Staubli VAL3: log.dtx

num nIndex = 14
num nLogType[300]
  [0] = 2
  [1] = 2
  [2] = 2
  [3] = 2
  [4] = 2
  [5] = 2
  [6] = 2
  [7] = 2
  [8] = 2
  [9] = 2
  [10] = 2
  [11] = 2
  [12] = 3
  [13] = 1
  [14] = 2
  [15] = 2
  [16] = 1
  [17] = 3
  [18] = 3
  [19] = 1
  [20] = 3
  [21] = 1
  [22] = 2
  [23] = 3
  [24] = 2
  [25] = 3
  [26] = 3
  [27] = 2
  [28] = 2
  [29] = 2
  [30] = 3
  [31] = 3
  [32] = 3
  [33] = 3
  [34] = 3
  [35] = 3
  [36] = 3
  [37] = 3
  [38] = 3
  [39] = 3
  [40] = 1
  [41] = 3
  [42] = 1
  [43] = 3
  [44] = 1
  [45] = 2
  [46] = 3
  [47] = 2
  [48] = 3
  [49] = 3
  [50] = 2
  [51] = 3
  [52] = 2
  [53] = 1
  [54] = 3
  [55] = 1
  [56] = 3
  [57] = 1
  [58] = 3
  [59] = 1
  [60] = 3
  [61] = 1
  [62] = 3
  [63] = 1
  [64] = 1
  [65] = 3
  [66] = 3
  [67] = 3
  [68] = 3
  [69] = 3
  [70] = 3
  [71] = 3
  [72] = 3
  [73] = 3
  [74] = 3
  [75] = 1
  [76] = 3
  [77] = 1
  [78] = 3
  [79] = 1
  [80] = 2
  [81] = 3
  [82] = 2
  [83] = 3
  [84] = 3
  [85] = 2
  [86] = 3
  [87] = 3
  [88] = 3
  [89] = 3
  [90] = 3
  [91] = 1
  [92] = 3
  [93] = 3
  [94] = 3
  [95] = 1
  [96] = 2
  [97] = 3
  [98] = 3
  [99] = 2
  [100] = 3
  [101] = 3
  [102] = 3
  [103] = 3
  [104] = 3
  [105] = 3
  [106] = 3
  [107] = 3
  [108] = 3
  [109] = 3
  [110] = 3
  [111] = 3
  [112] = 3
  [113] = 1
  [114] = 3
  [115] = 1
  [116] = 3
  [117] = 3
  [118] = 1
  [119] = 2
  [120] = 3
  [121] = 2
  [122] = 2
  [123] = 2
  [124] = 3
  [125] = 3
  [126] = 3
  [127] = 3
  [128] = 3
  [129] = 2
  [130] = 3
  [131] = 2
  [132] = 3
  [133] = 2
  [134] = 3
  [135] = 2
  [136] = 3
  [137] = 2
  [138] = 3
  [139] = 2
  [140] = 3
  [141] = 2
  [142] = 3
  [143] = 3
  [144] = 2
  [145] = 2
  [146] = 2
  [147] = 2
  [148] = 2
  [149] = 2
  [150] = 2
  [151] = 2
  [152] = 2
  [153] = 2
  [154] = 2
  [155] = 2
  [156] = 2
  [157] = 2
  [158] = 2
  [159] = 2
  [160] = 2
  [161] = 2
  [162] = 2
  [163] = 2
  [164] = 2
  [165] = 2
  [166] = 2
  [167] = 2
  [168] = 2
  [169] = 2
  [170] = 2
  [171] = 2
  [172] = 2
  [173] = 2
  [174] = 2
  [175] = 2
  [176] = 2
  [177] = 2
  [178] = 2
  [179] = 2
  [180] = 1
  [181] = 3
  [182] = 3
  [183] = 3
  [184] = 1
  [185] = 3
  [186] = 3
  [187] = 1
  [188] = 3
  [189] = 2
  [190] = 3
  [191] = 3
  [192] = 3
  [193] = 3
  [194] = 3
  [195] = 2
  [196] = 3
  [197] = 3
  [198] = 3
  [199] = 3
  [200] = 3
  [201] = 3
  [202] = 1
  [203] = 3
  [204] = 3
  [205] = 3
  [206] = 3
  [207] = 1
  [208] = 3
  [209] = 3
  [210] = 1
  [211] = 2
  [212] = 3
  [213] = 2
  [214] = 2
  [215] = 2
  [216] = 3
  [217] = 3
  [218] = 2
  [219] = 2
  [220] = 3
  [221] = 3
  [222] = 2
  [223] = 2
  [224] = 3
  [225] = 2
  [226] = 3
  [227] = 2
  [228] = 3
  [229] = 2
  [230] = 3
  [231] = 3
  [232] = 2
  [233] = 2
  [234] = 2
  [235] = 2
  [236] = 2
  [237] = 2
  [238] = 2
  [239] = 2
  [240] = 2
  [241] = 2
  [242] = 2
  [243] = 2
  [244] = 2
  [245] = 2
  [246] = 2
  [247] = 2
  [248] = 2
  [249] = 2
  [250] = 1
  [251] = 3
  [252] = 3
  [253] = 3
  [254] = 1
  [255] = 3
  [256] = 3
  [257] = 3
  [258] = 1
  [259] = 2
  [260] = 3
  [261] = 3
  [262] = 3
  [263] = 2
  [264] = 3
  [265] = 3
  [266] = 1
  [267] = 3
  [268] = 3
  [269] = 1
  [270] = 3
  [271] = 1
  [272] = 2
  [273] = 3
  [274] = 2
  [275] = 2
  [276] = 3
  [277] = 2
  [278] = 2
  [279] = 3
  [280] = 2
  [281] = 2
  [282] = 3
  [283] = 2
  [284] = 3
  [285] = 2
  [286] = 3
  [287] = 2
  [288] = 3
  [289] = 2
  [290] = 3
  [291] = 3
  [292] = 2
  [293] = 2
  [294] = 2
  [295] = 2
  [296] = 2
  [297] = 2
  [298] = 2
  [299] = 2
string sLog[300]
  [0] = "258.828 [路径信息]:移动到:12, L[271,-458,568,-7,-3,28]_spd=100%_b=50 09-16 10:48:04"
  [1] = "258.944 [路径信息]:移动到:13, L[271,-423,568,-7,-3,28]_spd=100%_b=50 09-16 10:48:04"
  [2] = "259.064 [路径信息]:移动到:14, L[241,-401,568,-7,-3,28]_spd=100%_b=50 09-16 10:48:05"
  [3] = "259.184 [路径信息]:移动到:15, L[189,-422,568,-7,-3,28]_spd=100%_b=50 09-16 10:48:05"
  [4] = "259.328 [路径信息]:移动到:16, L[189,-458,568,-7,-3,28]_spd=100%_b=50 09-16 10:48:05"
  [5] = "259.444 [路径信息]:移动到:17, L[159,-434,568,-7,-3,28]_spd=100%_b=50 09-16 10:48:05"
  [6] = "259.564 [路径信息]:移动到:18, L[121,-459,568,-7,-3,28]_spd=100%_b=50 09-16 10:48:06"
  [7] = "259.684 [路径信息]:移动到:19, L[121,-424,568,-7,-3,28]_spd=100%_b=50 09-16 10:48:06"
  [8] = "259.804 [路径信息]:移动到:20, L[90,-399,568,-7,-3,28]_spd=100%_b=50 09-16 10:48:06"
  [9] = "259.944 [路径信息]:移动到:21, L[40,-417,568,-7,-3,28]_spd=100%_b=50 09-16 10:48:06"
  [10] = "260.092 [路径信息]:移动到:22, L[40,-456,568,-7,-3,28]_spd=100%_b=50 09-16 10:48:07"
  [11] = "260.184 [路径信息]:移动到:23, L[3,-425,568,-7,-3,28]_spd=100%_b=50 09-16 10:48:07"
  [12] = "260.184 [信号信息]:dOut6=OFF 09-16 10:48:07"
  [13] = "261.184 [状态信息]:错误：-303. :0自动运行过程中伺服异常下电 09-16 10:48:09"
  [14] = "1112.913 [路径信息]:移动到:2, DOUT[70]-备用=TRUE 07-21 20:12:43"
  [15] = "1112.94  [路径信息]:移动到:3, wait->DIN[70]-备用=TRUE 07-21 20:12:43"
  [16] = "1294.838 [状态信息]:页面设置复位信号 07-21 20:17:28"
  [17] = "1297.928 [信号信息]:dOut10=OFF 07-21 20:17:33"
  [18] = "1298.8   [信号信息]:dOut6=ON 07-21 20:17:35"
  [19] = "1299.434 [状态信息]:程序号:1,J1MaxForce：0   ,J2MaxForce：152.6 ,J3MaxForce：73   ,J4MaxForce：1.3 ,J5MaxForce：10.03,J6MaxForce：0    07-21 20:17:36"
  [20] = "1299.434 [信号信息]:dOut1=ON 07-21 20:17:36"
  [21] = "1306.503 [状态信息]:当前处于生产状态 07-21 20:17:47"
  [22] = "1306.503 [路径信息]:移动到:0, DELAY = 1     s 07-21 20:17:47"
  [23] = "1306.503 [信号信息]:dOut2=ON 07-21 20:17:47"
  [24] = "1307.526 [路径信息]:移动到:1, L[1169,127,-142,15,129,-19]_spd=100%_b=0 07-21 20:17:48"
  [25] = "1307.526 [信号信息]:dOut8=ON 07-21 20:17:48"
  [26] = "1309.081 [信号信息]:dOut5=OFF 07-21 20:17:51"
  [27] = "1311.831 [路径信息]:移动到:2, L[1169,266,-142,15,129,-19]_spd=100%_b=0 07-21 20:17:55"
  [28] = "1316.763 [路径信息]:移动到轨迹PR01Washing001:3, WASH_DELAY = 0     s 07-21 20:18:03"
  [29] = "1316.784 [路径信息]:移动到:4, L[1169,266,-142,26,129,-19]_spd=100%_b=0 07-21 20:18:03"
  [30] = "1321.135 [信号信息]:dOut6=OFF 07-21 20:18:10"
  [31] = "180.317 [信号信息]:dOut97=ON 07-21 20:48:43"
  [32] = "196.059 [信号信息]:dOut6=ON 07-21 20:49:08"
  [33] = "196.677 [信号信息]:dOut8=ON 07-21 20:49:09"
  [34] = "197.418 [信号信息]:dOut97=OFF 07-21 20:49:10"
  [35] = "198.018 [信号信息]:dOut8=OFF 07-21 20:49:11"
  [36] = "199.801 [信号信息]:dOut8=ON 07-21 20:49:14"
  [37] = "203.867 [信号信息]:dOut5=ON 07-21 20:49:20"
  [38] = "204.256 [信号信息]:dOut8=OFF 07-21 20:49:21"
  [39] = "208.562 [信号信息]:dOut10=OFF 07-21 20:49:28"
  [40] = "212.136 [状态信息]:页面设置复位信号 07-21 20:49:33"
  [41] = "213.265 [信号信息]:dOut6=ON 07-21 20:49:35"
  [42] = "213.865 [状态信息]:当前处于ready状态 07-21 20:49:36"
  [43] = "213.887 [信号信息]:dOut1=ON 07-21 20:49:36"
  [44] = "251.032 [状态信息]:当前处于生产状态 07-21 20:50:34"
  [45] = "251.032 [路径信息]:移动到:0, DELAY = 1     s 07-21 20:50:34"
  [46] = "251.032 [信号信息]:dOut2=ON 07-21 20:50:34"
  [47] = "252.064 [路径信息]:移动到:1, L[1169,127,-142,15,129,-19]_spd=100%_b=0 07-21 20:50:36"
  [48] = "252.064 [信号信息]:dOut8=ON 07-21 20:50:36"
  [49] = "253.63  [信号信息]:dOut5=OFF 07-21 20:50:38"
  [50] = "256.347 [路径信息]:移动到:2, L[1169,266,-142,15,129,-19]_spd=100%_b=0 07-21 20:50:42"
  [51] = "261.222 [信号信息]:dOut6=OFF 07-21 20:50:50"
  [52] = "261.284 [路径信息]:移动到:4, L[1169,266,-142,26,129,-19]_spd=100%_b=0 07-21 20:50:50"
  [53] = "262.212 [状态信息]:错误：-303. :0自动运行过程中伺服异常下电 07-21 20:50:52"
  [54] = "262.733 [信号信息]:dOut11=ON 07-21 20:50:52"
  [55] = "262.759 [状态信息]:当前处于暂停状态 07-21 20:50:52"
  [56] = "262.759 [信号信息]:dOut3=ON 07-21 20:50:52"
  [57] = "264.227 [状态信息]:当前处于生产停止状态 07-21 20:50:55"
  [58] = "264.227 [信号信息]:dOut0=ON 07-21 20:50:55"
  [59] = "269.89  [状态信息]:收到页面点击清除报错! 07-21 20:51:04"
  [60] = "269.915 [信号信息]:dOut11=OFF 07-21 20:51:04"
  [61] = "273.022 [状态信息]:收到页面手动路径回Home点信号 07-21 20:51:09"
  [62] = "276.855 [信号信息]:dOut6=ON 07-21 20:51:15"
  [63] = "299.325 [状态信息]:页面设置复位信号 07-21 20:51:50"
  [64] = "301.959 [状态信息]:收到页面手动路径回Home点信号 07-21 20:51:54"
  [65] = "565.227 [信号信息]:dOut8=ON 07-21 20:58:47"
  [66] = "567.33  [信号信息]:dOut8=OFF 07-21 20:58:50"
  [67] = "571.862 [信号信息]:dOut8=ON 07-21 20:58:57"
  [68] = "572.394 [信号信息]:dOut8=OFF 07-21 20:58:58"
  [69] = "572.469 [信号信息]:dOut8=ON 07-21 20:58:58"
  [70] = "573.584 [信号信息]:dOut8=OFF 07-21 20:59:00"
  [71] = "575.243 [信号信息]:dOut8=ON 07-21 20:59:02"
  [72] = "575.802 [信号信息]:dOut5=ON 07-21 20:59:03"
  [73] = "576.029 [信号信息]:dOut8=OFF 07-21 20:59:04"
  [74] = "589.435 [信号信息]:dOut10=OFF 07-21 20:59:25"
  [75] = "604.459 [状态信息]:页面设置复位信号 07-21 20:59:48"
  [76] = "605.601 [信号信息]:dOut6=ON 07-21 20:59:50"
  [77] = "606.232 [状态信息]:程序号:1,J1MaxForce：67.45,J2MaxForce：264.18,J3MaxForce：102.39,J4MaxForce：8.71,J5MaxForce：19.2 ,J6MaxForce：1.88 07-21 20:59:51"
  [78] = "606.232 [信号信息]:dOut1=ON 07-21 20:59:51"
  [79] = "612.58  [状态信息]:当前处于生产状态 07-21 21:00:01"
  [80] = "612.58  [路径信息]:移动到:0, DELAY = 1     s 07-21 21:00:01"
  [81] = "612.58  [信号信息]:dOut2=ON 07-21 21:00:01"
  [82] = "613.621 [路径信息]:移动到:1, L[1169,127,-142,15,129,-19]_spd=100%_b=0 07-21 21:00:02"
  [83] = "613.621 [信号信息]:dOut8=ON 07-21 21:00:02"
  [84] = "615.161 [信号信息]:dOut5=OFF 07-21 21:00:05"
  [85] = "617.895 [路径信息]:移动到:2, L[1169,266,-142,15,129,-19]_spd=100%_b=0 07-21 21:00:09"
  [86] = "620.296 [信号信息]:dOut8=OFF 07-21 21:00:13"
  [87] = "620.788 [信号信息]:dOut6=OFF 07-21 21:00:14"
  [88] = "9.52  [信号信息]:dOut10=ON 09-16 10:39:57"
  [89] = "19.528 [信号信息]:dOut10=OFF 09-16 10:40:17"
  [90] = "60.184 [信号信息]:dIn0=ON 09-16 10:41:36"
  [91] = "60.312 [状态信息]:收到PLC复位信号 09-16 10:41:37"
  [92] = "60.828 [信号信息]:dIn0=OFF 09-16 10:41:38"
  [93] = "61.828 [信号信息]:dOut6=ON 09-16 10:41:40"
  [94] = "67.68  [信号信息]:dIn9=ON 09-16 10:41:51"
  [95] = "67.704 [状态信息]:收到PLC直接回Home点信号 09-16 10:41:51"
  [96] = "67.704 [路径信息]:直接回原点过程中 09-16 10:41:51"
  [97] = "67.704 [信号信息]:dOut8=ON 09-16 10:41:51"
  [98] = "68.564 [信号信息]:dOut5=ON 09-16 10:41:53"
  [99] = "68.796 [路径信息]:直接回原点完成 09-16 10:41:53"
  [100] = "68.796 [信号信息]:dOut6=OFF 09-16 10:41:53"
  [101] = "68.844 [信号信息]:dOut8=OFF 09-16 10:41:53"
  [102] = "69.076 [信号信息]:dOut0=ON 09-16 10:41:54"
  [103] = "69.404 [信号信息]:dIn9=OFF 09-16 10:41:54"
  [104] = "73.4   [信号信息]:dIn1=ON 09-16 10:42:02"
  [105] = "74.62  [信号信息]:dIn1=OFF 09-16 10:42:05"
  [106] = "87.112 [信号信息]:dOut8=ON 09-16 10:42:29"
  [107] = "87.18  [信号信息]:dOut8=OFF 09-16 10:42:29"
  [108] = "88.984 [信号信息]:dIn1=ON 09-16 10:42:33"
  [109] = "89.924 [信号信息]:dIn1=OFF 09-16 10:42:34"
  [110] = "102.18  [信号信息]:dIn1=ON 09-16 10:42:58"
  [111] = "109.252 [信号信息]:dIn1=OFF 09-16 10:43:12"
  [112] = "110.004 [信号信息]:dIn0=ON 09-16 10:43:14"
  [113] = "110.132 [状态信息]:收到PLC复位信号 09-16 10:43:14"
  [114] = "111.18  [信号信息]:dIn0=OFF 09-16 10:43:16"
  [115] = "112.78  [状态信息]:当前处于ready状态 09-16 10:43:19"
  [116] = "112.78  [信号信息]:dOut1=ON 09-16 10:43:19"
  [117] = "113.112 [信号信息]:dIn1=ON 09-16 10:43:20"
  [118] = "113.24  [状态信息]:当前处于生产状态 09-16 10:43:20"
  [119] = "113.24  [路径信息]:移动到:4, AOUT[4]-备用=0     09-16 10:43:20"
  [120] = "113.24  [信号信息]:dOut2=ON 09-16 10:43:20"
  [121] = "113.264 [路径信息]:移动到:10, DOUT[43]-吹干阀1=FALSE 09-16 10:43:20"
  [122] = "113.284 [路径信息]:移动到:14, DOUT[51]-吹干工作完成=FALSE 09-16 10:43:20"
  [123] = "113.308 [路径信息]:移动到:1, wait->DIN[20]-工作允许=TRUE 09-16 10:43:20"
  [124] = "114.424 [信号信息]:dIn1=OFF 09-16 10:43:22"
  [125] = "121.784 [信号信息]:dIn21=ON 09-16 10:43:37"
  [126] = "122.6   [信号信息]:dIn21=OFF 09-16 10:43:38"
  [127] = "125.18  [信号信息]:dIn40=ON 09-16 10:43:43"
  [128] = "125.82  [信号信息]:dIn40=OFF 09-16 10:43:45"
  [129] = "136.164 [路径信息]:移动到:0, DOUT[5]-机械人在home点=TRUE 09-16 10:44:05"
  [130] = "136.164 [信号信息]:dIn20=ON 09-16 10:44:05"
  [131] = "136.188 [路径信息]:移动到:2, DELAY = 0.5   s 09-16 10:44:05"
  [132] = "136.188 [信号信息]:dOut40=ON 09-16 10:44:05"
  [133] = "136.7   [路径信息]:移动到:3, wait->DIN[40]-私服位置到达=TRUE 09-16 10:44:06"
  [134] = "137.044 [信号信息]:dIn20=OFF 09-16 10:44:06"
  [135] = "138.724 [路径信息]:移动到:4, DELAY = 0.5   s 09-16 10:44:10"
  [136] = "138.724 [信号信息]:dIn40=ON 09-16 10:44:10"
  [137] = "139.232 [路径信息]:移动到:5, DOUT[40]-伺服旋转命令=FALSE 09-16 10:44:11"
  [138] = "139.232 [信号信息]:dOut40=OFF 09-16 10:44:11"
  [139] = "139.252 [路径信息]:移动到:2, L[61,-652,350,-2,-2,28]_spd=100%_b=50 09-16 10:44:11"
  [140] = "139.252 [信号信息]:dOut8=ON 09-16 10:44:11"
  [141] = "139.276 [路径信息]:移动到:3, L[489,-419,568,-7,-3,28]_spd=100%_b=50 09-16 10:44:11"
  [142] = "139.42  [信号信息]:dOut5=OFF 09-16 10:44:11"
  [143] = "139.744 [信号信息]:dIn40=OFF 09-16 10:44:12"
  [144] = "139.788 [路径信息]:移动到:4, L[489,-457,568,-7,-3,28]_spd=100%_b=50 09-16 10:44:12"
  [145] = "139.884 [路径信息]:移动到:5, L[459,-434,568,-7,-3,28]_spd=100%_b=50 09-16 10:44:12"
  [146] = "140.02  [路径信息]:移动到:6, L[427,-421,568,-7,-3,28]_spd=100%_b=50 09-16 10:44:12"
  [147] = "140.14  [路径信息]:移动到:7, L[427,-458,568,-7,-3,28]_spd=100%_b=50 09-16 10:44:12"
  [148] = "140.252 [路径信息]:移动到:8, L[393,-403,568,-7,-3,28]_spd=100%_b=50 09-16 10:44:13"
  [149] = "140.42  [路径信息]:移动到:9, L[345,-458,568,-7,-3,28]_spd=100%_b=50 09-16 10:44:13"
  [150] = "140.532 [路径信息]:移动到:10, L[345,-422,568,-7,-3,28]_spd=100%_b=50 09-16 10:44:13"
  [151] = "140.676 [路径信息]:移动到:11, L[312,-431,568,-7,-3,28]_spd=100%_b=50 09-16 10:44:14"
  [152] = "140.788 [路径信息]:移动到:12, L[271,-458,568,-7,-3,28]_spd=100%_b=50 09-16 10:44:14"
  [153] = "140.908 [路径信息]:移动到:13, L[271,-423,568,-7,-3,28]_spd=100%_b=50 09-16 10:44:14"
  [154] = "141.02  [路径信息]:移动到:14, L[241,-401,568,-7,-3,28]_spd=100%_b=50 09-16 10:44:14"
  [155] = "141.164 [路径信息]:移动到:15, L[189,-422,568,-7,-3,28]_spd=100%_b=50 09-16 10:44:14"
  [156] = "141.3   [路径信息]:移动到:16, L[189,-458,568,-7,-3,28]_spd=100%_b=50 09-16 10:44:15"
  [157] = "141.396 [路径信息]:移动到:17, L[159,-434,568,-7,-3,28]_spd=100%_b=50 09-16 10:44:15"
  [158] = "141.532 [路径信息]:移动到:18, L[121,-459,568,-7,-3,28]_spd=100%_b=50 09-16 10:44:15"
  [159] = "141.652 [路径信息]:移动到:19, L[121,-424,568,-7,-3,28]_spd=100%_b=50 09-16 10:44:15"
  [160] = "141.768 [路径信息]:移动到:20, L[90,-399,568,-7,-3,28]_spd=100%_b=50 09-16 10:44:16"
  [161] = "141.908 [路径信息]:移动到:21, L[40,-417,568,-7,-3,28]_spd=100%_b=50 09-16 10:44:16"
  [162] = "142.044 [路径信息]:移动到:22, L[40,-456,568,-7,-3,28]_spd=100%_b=50 09-16 10:44:16"
  [163] = "142.14  [路径信息]:移动到:23, L[3,-425,568,-7,-3,28]_spd=100%_b=50 09-16 10:44:16"
  [164] = "142.276 [路径信息]:移动到:24, L[-30,-459,568,-7,-3,28]_spd=100%_b=50 09-16 10:44:17"
  [165] = "142.396 [路径信息]:移动到:25, L[-30,-424,568,-7,-3,28]_spd=100%_b=50 09-16 10:44:17"
  [166] = "142.532 [路径信息]:移动到:26, L[-63,-402,568,-7,-3,28]_spd=100%_b=50 09-16 10:44:17"
  [167] = "142.652 [路径信息]:移动到:27, L[-112,-422,568,-7,-3,28]_spd=100%_b=50 09-16 10:44:17"
  [168] = "142.788 [路径信息]:移动到:28, L[-112,-459,568,-7,-3,28]_spd=100%_b=50 09-16 10:44:18"
  [169] = "142.908 [路径信息]:移动到:29, L[-149,-435,568,-7,-3,28]_spd=100%_b=50 09-16 10:44:18"
  [170] = "143.024 [路径信息]:移动到:30, L[-182,-460,568,-7,-3,28]_spd=100%_b=50 09-16 10:44:18"
  [171] = "143.14  [路径信息]:移动到:31, L[-182,-422,568,-7,-3,28]_spd=100%_b=50 09-16 10:44:18"
  [172] = "143.276 [路径信息]:移动到:32, L[-219,-406,568,-7,-3,28]_spd=100%_b=50 09-16 10:44:19"
  [173] = "143.42  [路径信息]:移动到:33, L[-267,-419,568,-7,-3,28]_spd=100%_b=50 09-16 10:44:19"
  [174] = "143.532 [路径信息]:移动到:34, L[-267,-457,568,-7,-3,28]_spd=100%_b=50 09-16 10:44:19"
  [175] = "143.676 [路径信息]:移动到:35, L[-308,-435,568,-7,-3,28]_spd=100%_b=50 09-16 10:44:19"
  [176] = "143.788 [路径信息]:移动到:36, L[-339,-459,568,-7,-3,28]_spd=100%_b=50 09-16 10:44:20"
  [177] = "143.908 [路径信息]:移动到:37, L[-339,-419,568,-7,-3,28]_spd=100%_b=50 09-16 10:44:20"
  [178] = "144.068 [路径信息]:移动到:38, L[-376,-400,568,-7,-3,28]_spd=100%_b=50 09-16 10:44:20"
  [179] = "144.164 [路径信息]:移动到:39, L[-338,-600,568,-7,-3,28]_spd=100%_b=50 09-16 10:44:20"
  [180] = "144.324 [状态信息]:页面设置停止信号 09-16 10:44:21"
  [181] = "144.324 [信号信息]:dOut2=OFF 09-16 10:44:21"
  [182] = "144.488 [信号信息]:dOut6=OFF 09-16 10:44:21"
  [183] = "144.556 [信号信息]:dOut8=OFF 09-16 10:44:21"
  [184] = "144.764 [状态信息]:当前处于生产停止状态 09-16 10:44:22"
  [185] = "144.764 [信号信息]:dOut42=OFF 09-16 10:44:22"
  [186] = "146.42  [信号信息]:dOut10=ON 09-16 10:44:25"
  [187] = "148.444 [状态信息]:收到页面手动路径回Home点信号 09-16 10:44:29"
  [188] = "150.532 [信号信息]:dOut6=ON 09-16 10:44:33"
  [189] = "151.724 [路径信息]:路径回原点过程中 09-16 10:44:35"
  [190] = "151.724 [信号信息]:dOut0=OFF 09-16 10:44:35"
  [191] = "154.7   [信号信息]:dOut8=ON 09-16 10:44:41"
  [192] = "179.3   [信号信息]:dOut8=OFF 09-16 10:45:29"
  [193] = "181.628 [信号信息]:dOut8=ON 09-16 10:45:33"
  [194] = "184.512 [信号信息]:dOut5=ON 09-16 10:45:39"
  [195] = "185.02  [路径信息]:路径回原点完成 09-16 10:45:40"
  [196] = "185.02  [信号信息]:dOut6=OFF 09-16 10:45:40"
  [197] = "185.3   [信号信息]:dOut0=ON 09-16 10:45:41"
  [198] = "188.236 [信号信息]:dOut10=OFF 09-16 10:45:46"
  [199] = "193.532 [信号信息]:dIn1=ON 09-16 10:45:57"
  [200] = "194.908 [信号信息]:dIn1=OFF 09-16 10:45:59"
  [201] = "195.468 [信号信息]:dIn0=ON 09-16 10:46:00"
  [202] = "195.596 [状态信息]:收到PLC复位信号 09-16 10:46:01"
  [203] = "196.128 [信号信息]:dIn0=OFF 09-16 10:46:02"
  [204] = "196.456 [信号信息]:dIn1=ON 09-16 10:46:02"
  [205] = "197.128 [信号信息]:dOut6=ON 09-16 10:46:04"
  [206] = "197.48  [信号信息]:dIn1=OFF 09-16 10:46:04"
  [207] = "197.74  [状态信息]:当前处于ready状态 09-16 10:46:05"
  [208] = "197.74  [信号信息]:dOut1=ON 09-16 10:46:05"
  [209] = "205.512 [信号信息]:dIn1=ON 09-16 10:46:20"
  [210] = "205.64  [状态信息]:当前处于生产状态 09-16 10:46:20"
  [211] = "205.64  [路径信息]:移动到:4, AOUT[4]-备用=0     09-16 10:46:20"
  [212] = "205.64  [信号信息]:dOut2=ON 09-16 10:46:20"
  [213] = "205.664 [路径信息]:移动到:10, DOUT[43]-吹干阀1=FALSE 09-16 10:46:20"
  [214] = "205.688 [路径信息]:移动到:0, DOUT[5]-机械人在home点=TRUE 09-16 10:46:20"
  [215] = "205.712 [路径信息]:移动到:1, wait->DIN[20]-工作允许=TRUE 09-16 10:46:20"
  [216] = "206.384 [信号信息]:dIn1=OFF 09-16 10:46:22"
  [217] = "210.444 [信号信息]:dIn20=ON 09-16 10:46:30"
  [218] = "210.468 [路径信息]:移动到:0, DOUT[40]-伺服旋转命令=TRUE 09-16 10:46:30"
  [219] = "210.492 [路径信息]:移动到:2, DELAY = 0.5   s 09-16 10:46:30"
  [220] = "210.492 [信号信息]:dOut40=ON 09-16 10:46:30"
  [221] = "210.92  [信号信息]:dIn20=OFF 09-16 10:46:31"
  [222] = "210.992 [路径信息]:移动到:3, wait->DIN[40]-私服位置到达=TRUE 09-16 10:46:31"
  [223] = "212.944 [路径信息]:移动到:4, DELAY = 0.5   s 09-16 10:46:35"
  [224] = "212.944 [信号信息]:dIn40=ON 09-16 10:46:35"
  [225] = "213.444 [路径信息]:移动到:0, DOUT[41]-清洗阀1=TRUE 09-16 10:46:36"
  [226] = "213.444 [信号信息]:dOut40=OFF 09-16 10:46:36"
  [227] = "213.468 [路径信息]:移动到:2, L[61,-652,350,-2,-2,28]_spd=100%_b=50 09-16 10:46:36"
  [228] = "213.468 [信号信息]:dOut8=ON 09-16 10:46:36"
  [229] = "213.492 [路径信息]:移动到:3, L[489,-419,568,-7,-3,28]_spd=100%_b=50 09-16 10:46:36"
  [230] = "213.628 [信号信息]:dOut5=OFF 09-16 10:46:36"
  [231] = "213.86  [信号信息]:dIn40=OFF 09-16 10:46:36"
  [232] = "213.98  [路径信息]:移动到:4, L[489,-457,568,-7,-3,28]_spd=100%_b=50 09-16 10:46:37"
  [233] = "214.092 [路径信息]:移动到:5, L[459,-434,568,-7,-3,28]_spd=100%_b=50 09-16 10:46:37"
  [234] = "214.236 [路径信息]:移动到:6, L[427,-421,568,-7,-3,28]_spd=100%_b=50 09-16 10:46:37"
  [235] = "214.348 [路径信息]:移动到:7, L[427,-458,568,-7,-3,28]_spd=100%_b=50 09-16 10:46:37"
  [236] = "214.468 [路径信息]:移动到:8, L[393,-403,568,-7,-3,28]_spd=100%_b=50 09-16 10:46:38"
  [237] = "214.604 [路径信息]:移动到:9, L[345,-458,568,-7,-3,28]_spd=100%_b=50 09-16 10:46:38"
  [238] = "214.748 [路径信息]:移动到:10, L[345,-422,568,-7,-3,28]_spd=100%_b=50 09-16 10:46:38"
  [239] = "214.884 [路径信息]:移动到:11, L[312,-431,568,-7,-3,28]_spd=100%_b=50 09-16 10:46:38"
  [240] = "214.98  [路径信息]:移动到:12, L[271,-458,568,-7,-3,28]_spd=100%_b=50 09-16 10:46:39"
  [241] = "215.116 [路径信息]:移动到:13, L[271,-423,568,-7,-3,28]_spd=100%_b=50 09-16 10:46:39"
  [242] = "215.236 [路径信息]:移动到:14, L[241,-401,568,-7,-3,28]_spd=100%_b=50 09-16 10:46:39"
  [243] = "215.36  [路径信息]:移动到:15, L[189,-422,568,-7,-3,28]_spd=100%_b=50 09-16 10:46:39"
  [244] = "215.504 [路径信息]:移动到:16, L[189,-458,568,-7,-3,28]_spd=100%_b=50 09-16 10:46:40"
  [245] = "215.592 [路径信息]:移动到:17, L[159,-434,568,-7,-3,28]_spd=100%_b=50 09-16 10:46:40"
  [246] = "215.74  [路径信息]:移动到:18, L[121,-459,568,-7,-3,28]_spd=100%_b=50 09-16 10:46:40"
  [247] = "215.86  [路径信息]:移动到:19, L[121,-424,568,-7,-3,28]_spd=100%_b=50 09-16 10:46:40"
  [248] = "215.98  [路径信息]:移动到:20, L[90,-399,568,-7,-3,28]_spd=100%_b=50 09-16 10:46:41"
  [249] = "216.116 [路径信息]:移动到:21, L[40,-417,568,-7,-3,28]_spd=100%_b=50 09-16 10:46:41"
  [250] = "216.164 [状态信息]:页面设置生产结束信号 09-16 10:46:41"
  [251] = "216.164 [信号信息]:dOut2=OFF 09-16 10:46:41"
  [252] = "216.372 [信号信息]:dOut8=OFF 09-16 10:46:41"
  [253] = "216.396 [信号信息]:dOut6=OFF 09-16 10:46:41"
  [254] = "216.652 [状态信息]:当前处于停止状态 09-16 10:46:42"
  [255] = "216.652 [信号信息]:dOut0=ON 09-16 10:46:42"
  [256] = "219.836 [信号信息]:dOut10=ON 09-16 10:46:48"
  [257] = "221.236 [信号信息]:dOut6=ON 09-16 10:46:51"
  [258] = "223.676 [状态信息]:收到页面手动路径回Home点信号 09-16 10:46:56"
  [259] = "223.676 [路径信息]:路径回原点过程中 09-16 10:46:56"
  [260] = "223.676 [信号信息]:dOut0=OFF 09-16 10:46:56"
  [261] = "224.652 [信号信息]:dOut8=ON 09-16 10:46:57"
  [262] = "239.26  [信号信息]:dOut5=ON 09-16 10:47:26"
  [263] = "239.748 [路径信息]:路径回原点完成 09-16 10:47:27"
  [264] = "239.748 [信号信息]:dOut6=OFF 09-16 10:47:27"
  [265] = "240.028 [信号信息]:dOut0=ON 09-16 10:47:28"
  [266] = "243.96  [状态信息]:页面设置复位信号 09-16 10:47:35"
  [267] = "246.36  [信号信息]:dOut10=OFF 09-16 10:47:40"
  [268] = "247.236 [信号信息]:dOut6=ON 09-16 10:47:42"
  [269] = "247.86  [状态信息]:程序号:1,J1MaxForce：264.44,J2MaxForce：326.51,J3MaxForce：123.34,J4MaxForce：18.83,J5MaxForce：15.47,J6MaxForce：3.53 09-16 10:47:43"
  [270] = "247.86  [信号信息]:dOut1=ON 09-16 10:47:43"
  [271] = "250.24  [状态信息]:当前处于生产状态 09-16 10:47:47"
  [272] = "250.24  [路径信息]:移动到:3, AOUT[1]-反馈速度=0     09-16 10:47:47"
  [273] = "250.24  [信号信息]:dOut2=ON 09-16 10:47:47"
  [274] = "250.26  [路径信息]:移动到:8, DOUT[41]-清洗阀1=FALSE 09-16 10:47:48"
  [275] = "250.284 [路径信息]:移动到:14, DOUT[51]-吹干工作完成=FALSE 09-16 10:47:48"
  [276] = "250.284 [信号信息]:dOut42=OFF 09-16 10:47:48"
  [277] = "250.304 [路径信息]:移动到:1, wait->DIN[20]-工作允许=TRUE 09-16 10:47:48"
  [278] = "254.652 [路径信息]:移动到:1, AOUT[5]-伺服执行定位号=5     09-16 10:47:56"
  [279] = "254.652 [信号信息]:dOut40=ON 09-16 10:47:56"
  [280] = "254.676 [路径信息]:移动到:2, DELAY = 0.5   s 09-16 10:47:56"
  [281] = "255.164 [路径信息]:移动到:3, wait->DIN[40]-私服位置到达=TRUE 09-16 10:47:57"
  [282] = "255.212 [信号信息]:dIn20=OFF 09-16 10:47:57"
  [283] = "256.768 [路径信息]:移动到:4, DELAY = 0.5   s 09-16 10:48:00"
  [284] = "256.768 [信号信息]:dIn40=ON 09-16 10:48:00"
  [285] = "257.268 [路径信息]:移动到:0, DOUT[41]-清洗阀1=TRUE 09-16 10:48:01"
  [286] = "257.268 [信号信息]:dOut40=OFF 09-16 10:48:01"
  [287] = "257.292 [路径信息]:移动到:2, L[61,-652,350,-2,-2,28]_spd=100%_b=50 09-16 10:48:01"
  [288] = "257.292 [信号信息]:dOut8=ON 09-16 10:48:01"
  [289] = "257.316 [路径信息]:移动到:3, L[489,-419,568,-7,-3,28]_spd=100%_b=50 09-16 10:48:01"
  [290] = "257.364 [信号信息]:dIn40=OFF 09-16 10:48:01"
  [291] = "257.456 [信号信息]:dOut5=OFF 09-16 10:48:02"
  [292] = "257.816 [路径信息]:移动到:4, L[489,-457,568,-7,-3,28]_spd=100%_b=50 09-16 10:48:02"
  [293] = "257.94  [路径信息]:移动到:5, L[459,-434,568,-7,-3,28]_spd=100%_b=50 09-16 10:48:03"
  [294] = "258.06  [路径信息]:移动到:6, L[427,-421,568,-7,-3,28]_spd=100%_b=50 09-16 10:48:03"
  [295] = "258.18  [路径信息]:移动到:7, L[427,-458,568,-7,-3,28]_spd=100%_b=50 09-16 10:48:03"
  [296] = "258.3   [路径信息]:移动到:8, L[393,-403,568,-7,-3,28]_spd=100%_b=50 09-16 10:48:03"
  [297] = "258.444 [路径信息]:移动到:9, L[345,-458,568,-7,-3,28]_spd=100%_b=50 09-16 10:48:03"
  [298] = "258.564 [路径信息]:移动到:10, L[345,-422,568,-7,-3,28]_spd=100%_b=50 09-16 10:48:04"
  [299] = "258.708 [路径信息]:移动到:11, L[312,-431,568,-7,-3,28]_spd=100%_b=50 09-16 10:48:04"
